FUNCTION_BLOCK FB_CylinderPos_MoveAbsolut
(*

The function block used to starts positioning to an absolute target position. 

Constructor: 		Patryk Panylo
Company:			E. Riexinger GmbH
Date:				22.09.2015
Version:			1.00

Date:			Revision:		Who:				Comment

*)
VAR_INPUT
	(* Input variables / Eingang Variablen *)
	bEnable						:BOOL;			(* Function block enable *)
	bNoEStop					:BOOL;			(* No ermergency Stop / Keine Notaus *)
	bLightCurtainOK				:BOOL;			(* Light curtain ok / Freigabe Lichtschranke i.o *)
	bAirPressure				:BOOL;			(* Signal air pressure *)
	arbInBase					:ARRAY[1..ungGr05CylinderPosMaxNo] OF BOOL;
	arbInWork					:ARRAY[1..ungGr05CylinderPosMaxNo] OF BOOL;
	arbInError					:ARRAY[1..ungGr05CylinderPosMaxNo] OF BOOL;
	bExecute					:BOOL;			(* Execut the function block *)
	lrPosition					:LREAL;			(* Absolute target position *)
	lrPosOffset					:LREAL;					(* Position offset *)
	lrOriginShiftPos			:LREAL;					(* Origin shift position *)
	etDirection					:ET_MC_Direction;			(* Direction: -1 Negative, +1 Positive *)
	usnCodingType				:USINT;
END_VAR
VAR_OUTPUT
	(* Output variables / Ausgang Variablen *)
	lrActPosition				:LREAL;			(* Absolute actual position *)
	arbToBase					:ARRAY[1..ungGr05CylinderPosMaxNo] OF BOOL;
	arbToWork					:ARRAY[1..ungGr05CylinderPosMaxNo] OF BOOL;
	bDone						:BOOL;			(* Program done *)
	bBusy						:BOOL;			(* Program busy *)
	bError						:BOOL;			(* Error *)
	udnErrorNo					:UDINT;			(* Error number *)
	sErrorMsg					:STRING; 		(* Error message *)
END_VAR
VAR_IN_OUT
	(* Input Output variables / Ausgang Variablen *)

END_VAR
VAR
	(* Enummerations *)
	etMC_States					:ET_MC_States := ET_MC_States_eInit;

	(* Variables *)
	wSetCylinderPos				:WORD;			(* Set position of cylinder  *)
	wGetCylinderPos				:WORD;			(* Get position of cylinder  *)

	wCylinderPos				:WORD;

	nWatchdog					:INT;

	bFirstTime					:BOOL;
	(* References *)

	(* Interfaces *)

	(* Instances *)
	rtExecute					:R_TRIG;

END_VAR


wGetCylinderPos.0 := arbInBase[1];
wGetCylinderPos.1 := arbInWork[1];
wGetCylinderPos.2 := arbInBase[2];
wGetCylinderPos.3 := arbInWork[2];
wGetCylinderPos.4 := arbInBase[3];
wGetCylinderPos.5 := arbInWork[3];

lrActPosition := F_GetCylinderPos(wGetCylinderPos, lrPosOffset, lrOriginShiftPos, etDirection, usnCodingType);

IF NOT bEnable
THEN
	bDone := bExecute AND bBusy;		(* Program done *)
	bBusy := bExecute;                                  	(* Program not busy *)
	bError := FALSE;                                 	(* Program not error *)
	udnErrorNo := 0;                                 		(* Error number *)

	bFirstTime := FALSE;
	RETURN;
END_IF

IF NOT bFirstTime
THEN
	bDone := FALSE;                                	(* Program done *)
	bBusy := FALSE;                                 	(* Program not busy *)
	bError := FALSE;                                 	(* Program not error *)
	udnErrorNo := 0;                                 		(* Error number *)

	etMC_States := ET_MC_States_eInit;                      (* Next step *)

	bFirstTime := TRUE;
END_IF;

rtExecute(CLK := bExecute
			     AND bNoEStop
			     AND bLightCurtainOK
			     AND bAirPressure
);

IF rtExecute.Q
THEN
	etMC_States := ET_MC_States_eInit;                      (* Next step *)

ELSIF NOT bExecute
	    OR NOT bNoEStop
	    OR NOT bLightCurtainOK
	    OR NOT bAirPressure
THEN
	arbToBase[1] := FALSE;
	arbToWork[1] := FALSE;
	arbToBase[2] := FALSE;
	arbToWork[2] := FALSE;
	arbToBase[3] := FALSE;
	arbToWork[3] := FALSE;

END_IF;

CASE etMC_States OF

	ET_MC_States_eInit:
		bBusy := FALSE;                                    	(* Program not busy *)
		bError := FALSE;                         		(* Program not error *)
		udnErrorNo := 0;                         		(* Error number *)

		IF rtExecute.Q
		THEN
			nWatchdog := 0;
			bDone := FALSE;				(* Program done, in position *)
			bBusy := TRUE;				(* Program busy *)

			IF bNoEStop
			     AND bLightCurtainOK
			     AND bAirPressure
			THEN
				etMC_States := ET_MC_States_eRunning;			(* Next step *)

			ELSE
				udnErrorNo := 4;                     (* Error number *)

				etMC_States := ET_MC_States_eError;			(* Next step *)

			END_IF;
		END_IF;

	ET_MC_States_eRunning:
		wSetCylinderPos := F_SetCylinderPos(lrPosition, lrPosOffset, lrOriginShiftPos, etDirection, usnCodingType);

		arbToBase[1] := wSetCylinderPos.0;
		arbToWork[1] := wSetCylinderPos.1;
		arbToBase[2] := wSetCylinderPos.2;
		arbToWork[2] := wSetCylinderPos.3;
		arbToBase[3] := wSetCylinderPos.4;
		arbToWork[3] := wSetCylinderPos.5;

		etMC_States := ET_MC_States_eWaiting;			(* Next step *)

	ET_MC_States_eWaiting:
		wCylinderPos.0 := arbToBase[1];
		wCylinderPos.1 := arbToWork[1];
		wCylinderPos.2 := arbToBase[2];
		wCylinderPos.3 := arbToWork[2];
		wCylinderPos.4 := arbToBase[3];
		wCylinderPos.5 := arbToWork[3];
		
		lrPosition := F_GetCylinderPos(wCylinderPos, lrPosOffset, lrOriginShiftPos, etDirection, usnCodingType);

		IF lrPosition = lrActPosition
		THEN
			arbToBase[1] := FALSE;
			arbToWork[1] := FALSE;
			arbToBase[2] := FALSE;
			arbToWork[2] := FALSE;
			arbToBase[3] := FALSE;
			arbToWork[3] := FALSE;

			etMC_States := ET_MC_States_eDone;			(* Next step *)

		ELSIF arbInError[1]
			    OR arbInError[2]
			    OR arbInError[3]
		THEN
			arbToBase[1] := FALSE;
			arbToWork[1] := FALSE;
			arbToBase[2] := FALSE;
			arbToWork[2] := FALSE;
			arbToBase[3] := FALSE;
			arbToWork[3] := FALSE;

			etMC_States := ET_MC_States_eError;			(* Next step *)

		END_IF;

	ET_MC_States_eDone:
		nWatchdog := 0;
		bDone := TRUE;			(* Program done, in position *)
		bBusy := FALSE;			(* Program not busy *)

		etMC_States := ET_MC_States_eNotExecute;            (* Next step *)

	ET_MC_States_eError:
		nWatchdog := 0;
		bDone := FALSE;			(* Program done, in position *)
		bError := TRUE;			(* Program error *)   
		bBusy := FALSE;			(* Program not busy *)

        		etMC_States := ET_MC_States_eNotExecute;			(*Next step *)

	ET_MC_States_eNotExecute:
		IF NOT bExecute
		THEN
			bDone := FALSE;					(* Program done, in position *)
			bBusy := FALSE;                                 	(* Program not busy *)
			bError := FALSE;                     			(* Program not error *)
			udnErrorNo := 0;                     			(* Error number *)

			etMC_States := ET_MC_States_eInit;			(* Next step *)
		
		END_IF;
END_CASE;

END_FUNCTION_BLOCK

(* stored: Version 1.1.0.1, ProductVersion 3.1.4024.15
   POU FB_CylinderPos_MoveAbsolut: Id {1fc26971-3434-4e4c-a581-36e9e4178b55}, SpecialFunc None *)
